(* IEC 61131-3 sources: avi-aoi-management/scripts/ai-eval/ngau-nhien/lib/st-scl/mau-scl/st-ud9-ghi-dich-loai-bo/src, 2 files *)

(* ---- LoaiBoAOI.st ---- *)
FUNCTION_BLOCK "LoaiBoAOI"
{ S7_Optimized_Access := 'TRUE' }
VERSION : 0.1
   VAR_INPUT
      ENCODER : Bool;
      CO_SAN_PHAM : Bool;
      LOI_AOI : Bool;
      RESET : Bool;
      VI_TRI_GAT : Int;
      T_GAT : Time;
   END_VAR

   VAR_OUTPUT
      CAN_GAT : Bool;
      DEM_GAT : DInt;
      SO_O_LOI : Int;
   END_VAR

   VAR
      rtEnc : R_TRIG;
      tg : "ThanhGhiDich";
      xungGat : TP_TIME;
   END_VAR

   VAR_TEMP
      toi : Bool;
   END_VAR

   REGION Dich thanh ghi theo encoder
      #rtEnc(CLK := #ENCODER);
      #tg(DICH := #rtEnc.Q AND NOT #RESET, GHI := #CO_SAN_PHAM AND #LOI_AOI AND NOT #RESET, XOA := #RESET, VI_TRI := #VI_TRI_GAT);
      // sản phẩm lỗi vừa được dịch tới vị trí gạt
      #toi := #rtEnc.Q AND NOT #RESET AND #VI_TRI_GAT >= 1 AND #VI_TRI_GAT <= 32 AND #tg.Q;
   END_REGION

   REGION Dem va gat
      IF #RESET THEN
         #DEM_GAT := 0;
      ELSIF #toi THEN
         #DEM_GAT := #DEM_GAT + 1;
      END_IF;
      #xungGat(IN := #toi, PT := #T_GAT);
      #CAN_GAT := #xungGat.Q;
      #SO_O_LOI := #tg.SO_O;
   END_REGION
END_FUNCTION_BLOCK

(* ---- ThanhGhiDich.st ---- *)
FUNCTION_BLOCK "ThanhGhiDich"
{ S7_Optimized_Access := 'TRUE' }
VERSION : 0.1
   VAR_INPUT
      DICH : Bool;
      GHI : Bool;
      XOA : Bool;
      VI_TRI : Int;
   END_VAR

   VAR_OUTPUT
      Q : Bool;
      SO_O : Int;
   END_VAR

   VAR
      o : Array[0..32] of Bool;
   END_VAR

   VAR_TEMP
      i : Int;
   END_VAR

   REGION Cap nhat thanh ghi
      IF #XOA THEN
         FOR #i := 0 TO 32 DO #o[#i] := FALSE; END_FOR;
      ELSE
         IF #DICH THEN
            FOR #i := 32 TO 1 BY -1 DO #o[#i] := #o[#i - 1]; END_FOR;
            #o[0] := FALSE;
         END_IF;
         IF #GHI THEN
            #o[0] := TRUE;
         END_IF;
      END_IF;
   END_REGION

   REGION Doc vi tri va dem o
      IF #VI_TRI >= 0 AND #VI_TRI <= 32 THEN
         #Q := #o[#VI_TRI];
      ELSE
         #Q := FALSE;
      END_IF;
      #SO_O := 0;
      FOR #i := 0 TO 32 DO
         IF #o[#i] THEN #SO_O := #SO_O + 1; END_IF;
      END_FOR;
   END_REGION
END_FUNCTION_BLOCK
